(* IEC 61131-3 sources: codesys-framework/txt/application/WeVe Core (library)/60 Event/Service/FB_EventService/Properties, 3 files *)

(* ---- HasAlarm.prop.st ---- *)
PROPERTY HasAlarm : BOOL
// --- BEGIN IMPLEMENTATION ---

// ----------- GET -----------
VAR
END_VAR

// -- BEGIN IMPLEMENTATION GET --
HasAlarm := _scState.xAlarmIsOn;

(* ---- HasWarning.prop.st ---- *)
PROPERTY HasWarning : BOOL
// --- BEGIN IMPLEMENTATION ---

// ----------- GET -----------
VAR
END_VAR

// -- BEGIN IMPLEMENTATION GET --
HasWarning := _scState.xWarningIsOn;

(* ---- State.prop.st ---- *)
PROPERTY State : SC_EventState
// --- BEGIN IMPLEMENTATION ---

// ----------- GET -----------
VAR
END_VAR

// -- BEGIN IMPLEMENTATION GET --
State := _scState;
